// TIA Portal V21 export
Screen "TiaMcpLibraryScreen"  800x480, Number=1
